Universal Robots URScript: T001_openai_gpt-oss-120b_baseline_rep2.urscript

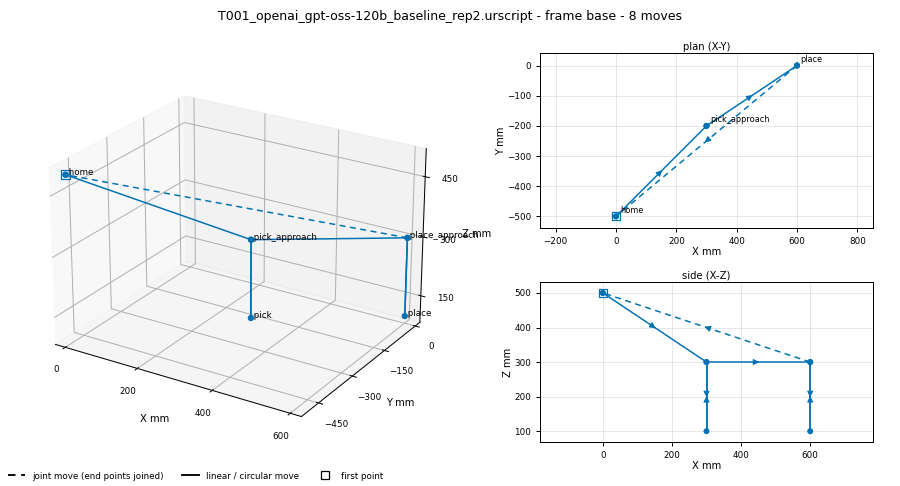
[picture p0: tool path of T001_openai_gpt-oss-120b_baseline_rep2.urscript in frame base, 8 of 8 moves have a stored position in this frame; points joined in program order, loops and branches not executed]
def main():
    # Payload configuration (mass in kg, CoG in meters)
    set_payload(0.5, 0.0, 0.0, 0.0, 0.0, 0.0)

    # TCP speed limit (max 250 mm/s = 0.25 m/s)
    set_tcp_speed(0.25)

    # -------------------------------------------------
    # Define key waypoints (positions in meters, orientation in radians)
    # -------------------------------------------------
    home            = p[0.0, -0.5, 0.5, 0, 3.14, 0]
    pick_approach   = p[0.30, -0.20, 0.30, 0, 3.14, 0]
    pick            = p[0.30, -0.20, 0.10, 0, 3.14, 0]
    lift            = p[0.30, -0.20, 0.30, 0, 3.14, 0]
    place_approach  = p[0.60,  0.00, 0.30, 0, 3.14, 0]
    place           = p[0.60,  0.00, 0.10, 0, 3.14, 0]
    retreat         = p[0.60,  0.00, 0.30, 0, 3.14, 0]

    # -------------------------------------------------
    # 1) Move to home position (joint move)
    # -------------------------------------------------
    movej(home, a=1.4, v=0.20, t=0, r=0)

    # -------------------------------------------------
    # 2) Approach pick point (linear move, 200 mm/s)
    # -------------------------------------------------
    movel(pick_approach, a=1.2, v=0.20, t=0, r=0)

    # -------------------------------------------------
    # 3) Descend to pick (linear move, 100 mm/s)
    # -------------------------------------------------
    movel(pick, a=1.0, v=0.10, t=0, r=0)

    # Gripper close (placeholder – replace with actual command)
    set_digital_out(8, True)

    # -------------------------------------------------
    # 4) Lift from pick (linear move, 150 mm/s)
    # -------------------------------------------------
    movel(lift, a=1.2, v=0.15, t=0, r=0)

    # -------------------------------------------------
    # 5) Transit to place approach (linear move, 200 mm/s)
    # -------------------------------------------------
    movel(place_approach, a=1.4, v=0.20, t=0, r=0)

    # -------------------------------------------------
    # 6) Descend to place (linear move, 100 mm/s)
    # -------------------------------------------------
    movel(place, a=1.0, v=0.10, t=0, r=0)

    # Gripper open (placeholder – replace with actual command)
    set_digital_out(8, False)

    # -------------------------------------------------
    # 7) Retreat from place (linear move, 150 mm/s)
    # -------------------------------------------------
    movel(retreat, a=1.2, v=0.15, t=0, r=0)

    # -------------------------------------------------
    # 8) Return to home position (joint move)
    # -------------------------------------------------
    movej(home, a=1.4, v=0.20, t=0, r=0)

end
